RESOURCE RES0 : EMB_RES_ECO
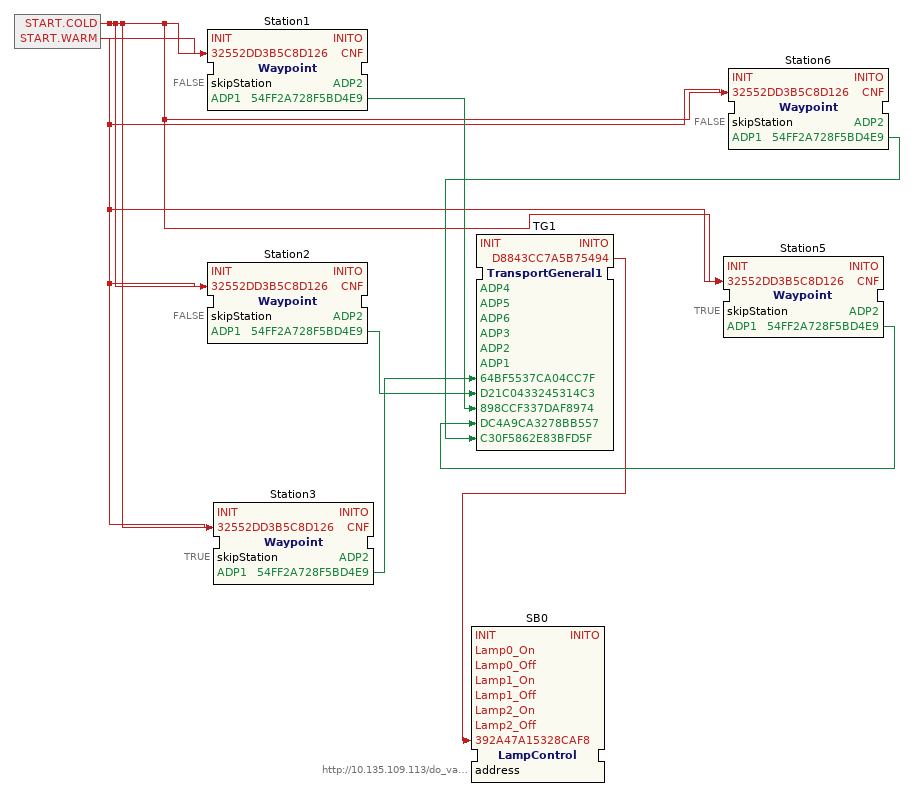
  FBS
    Station1 : Waypoint(skipStation := FALSE);
    Station2 : Waypoint(skipStation := FALSE);
    Station3 : Waypoint(skipStation := TRUE);
    TG1 : TransportGeneral1;
    SB0 : LampControl(address := http://10.135.109.113/do_value/slot_0);
    Station5 : Waypoint(skipStation := TRUE);
    Station6 : Waypoint(skipStation := FALSE);
  END_FBS
  EVENT_CONNECTIONS
    START.COLD TO Station2.32552DD3B5C8D126;
    START.COLD TO Station3.32552DD3B5C8D126;
    START.COLD TO Station5.32552DD3B5C8D126;
    START.COLD TO Station6.32552DD3B5C8D126;
    START.WARM TO Station2.32552DD3B5C8D126;
    START.WARM TO Station3.32552DD3B5C8D126;
    START.WARM TO Station5.32552DD3B5C8D126;
    START.WARM TO Station6.32552DD3B5C8D126;
    TG1.D8843CC7A5B75494 TO SB0.392A47A15328CAF8;
    START.COLD TO Station1.32552DD3B5C8D126;
    START.WARM TO Station1.32552DD3B5C8D126;
  END_CONNECTIONS
  ADAPTER_CONNECTIONS
    Station3.54FF2A728F5BD4E9 TO TG1.64BF5537CA04CC7F;
    Station2.54FF2A728F5BD4E9 TO TG1.D21C0433245314C3;
    Station1.54FF2A728F5BD4E9 TO TG1.898CCF337DAF8974;
    Station5.54FF2A728F5BD4E9 TO TG1.DC4A9CA3278BB557;
    Station6.54FF2A728F5BD4E9 TO TG1.C30F5862E83BFD5F;
  END_CONNECTIONS
END_RESOURCE
